PROGRAM main
  VAR
    S1 AT %IX0.0 : BOOL; (* barrera de entrada: entra un auto *)
    S2 AT %IX0.1 : BOOL; (* barrera de salida: sale un auto *)
    H1 AT %QX0.0 : BOOL; (* verde: hay lugar *)
    H2 AT %QX0.1 : BOOL; (* amarillo: lleno *)
    F_ENTRA      : R_TRIG;
    F_SALE       : R_TRIG;
    AUTOS        : INT; (* autos adentro *)
    LIBRES       : INT; (* lugares libres *)
    HAY_LUGAR    : BOOL; (* AUTOS < capacidad *)
    HAY_AUTOS    : BOOL; (* AUTOS > 0 *)
  END_VAR
  VAR  (* added by the conversion: wires and edge detectors of the diagram *)
    R_TRIG1 : R_TRIG;
    R_TRIG2 : R_TRIG;
  END_VAR

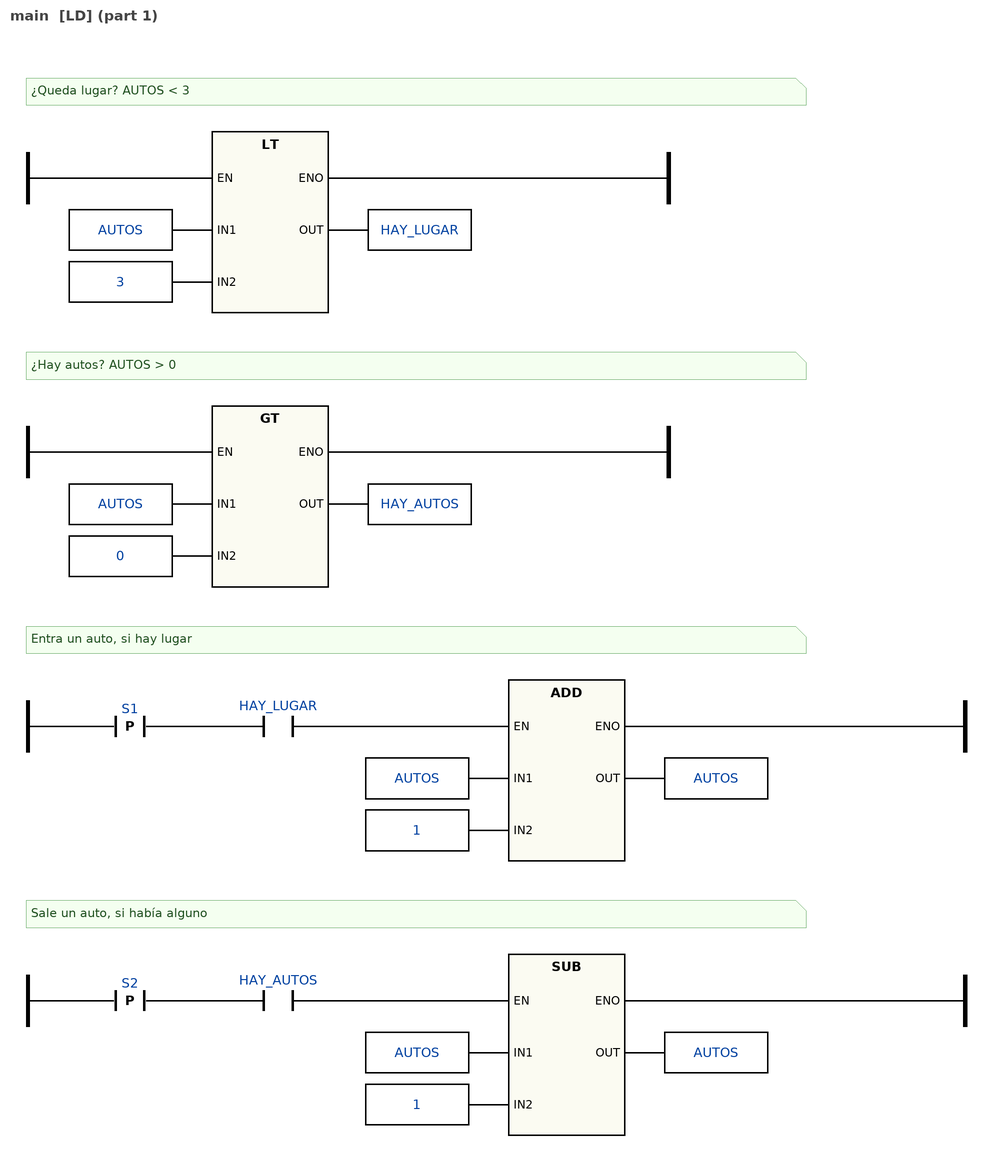
(* LD diagram, written out as Structured Text *)
(* ¿Queda lugar? AUTOS < 3 *)
HAY_LUGAR := AUTOS < 3;
(* ¿Hay autos? AUTOS > 0 *)
HAY_AUTOS := AUTOS > 0;
(* Entra un auto, si hay lugar *)
R_TRIG1(CLK := S1);
IF R_TRIG1.Q AND HAY_LUGAR THEN AUTOS := AUTOS + 1; END_IF;
(* Sale un auto, si había alguno *)
R_TRIG2(CLK := S2);
IF R_TRIG2.Q AND HAY_AUTOS THEN AUTOS := AUTOS - 1; END_IF;
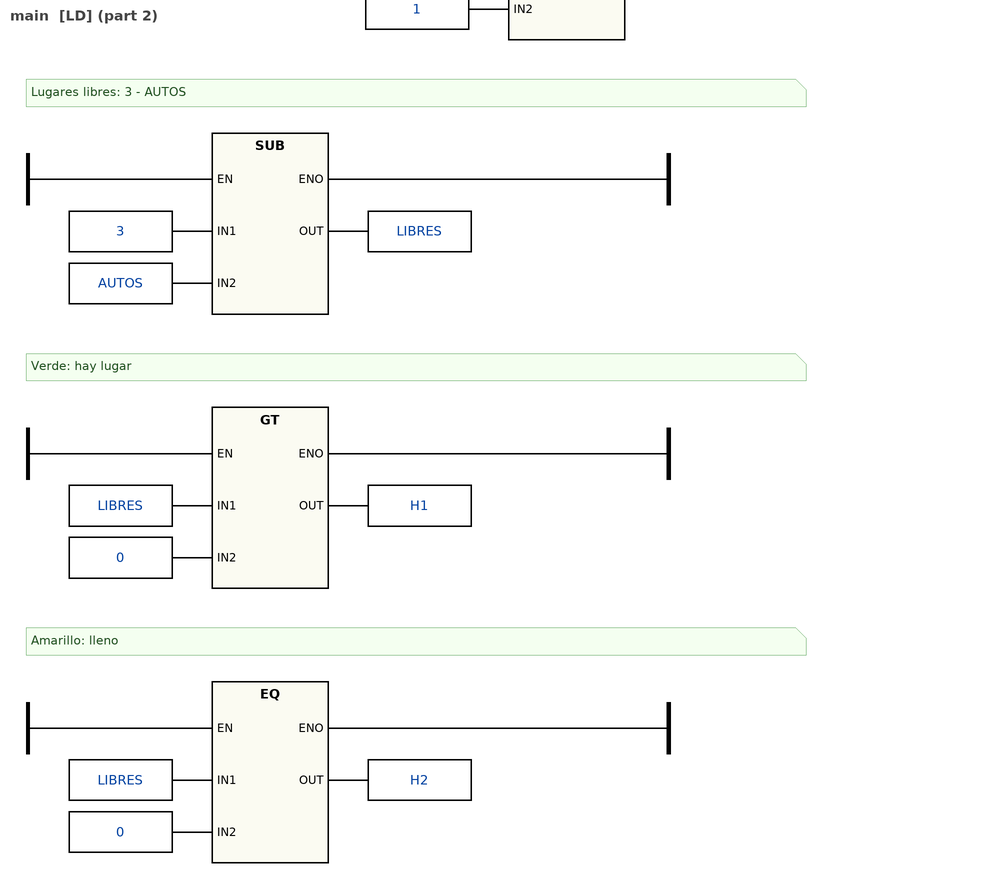
(* Lugares libres: 3 - AUTOS *)
LIBRES := 3 - AUTOS;
(* Verde: hay lugar *)
H1 := LIBRES > 0;
(* Amarillo: lleno *)
H2 := LIBRES = 0;
END_PROGRAM
